// LS Electric XG5000 project: Trafic light3T
// PLC NewPLC
// module base 0 slot 0: Input/Output Module:XBM-DN32S (DC 24V INPUT/TR OUTPUT, 32points)
// module base 0 slot 1: Analog Input Module:XBF-AD04A (Volt/Current, 4-CH)
// module base 0 slot 2: Analog Output Module:XBF-DV04A (Voltage, 4-CH)

PROGRAM NewProgram (task: Scan Program)

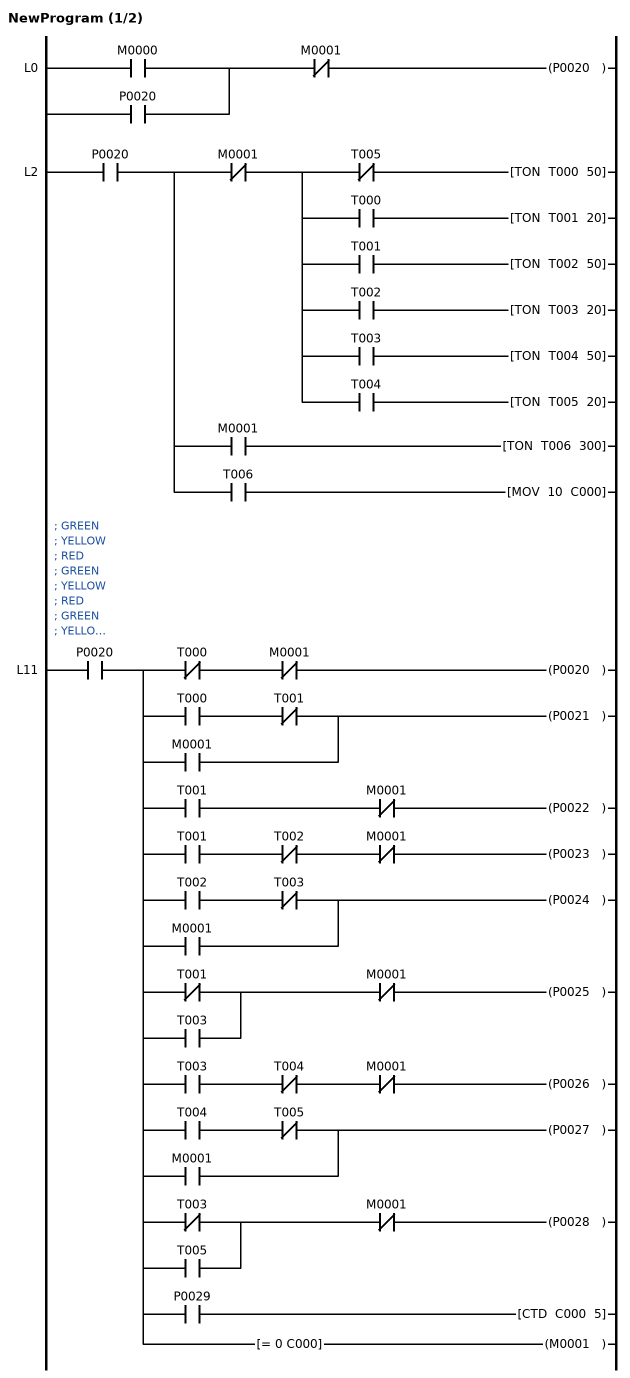
; L0
LOAD      M0000
OR        P0020
AND NOT   M0001
OUT       P0020
; L2
LOAD      P0020
MPUSH
AND NOT   M0001
MPUSH
AND NOT   T005
TON       T000 50
MLOAD
AND       T000
TON       T001 20
MLOAD
AND       T001
TON       T002 50
MLOAD
AND       T002
TON       T003 20
MLOAD
AND       T003
TON       T004 50
MPOP
AND       T004
TON       T005 20
MLOAD
AND       M0001
TON       T006 300
MPOP
AND       T006
MOV       10 C000
// output comment: 
; L11
LOAD      P0020
MPUSH
AND NOT   T000
AND NOT   M0001
OUT       P0020
MLOAD
LOAD      T000
AND NOT   T001
OR        M0001
AND LOAD
OUT       P0021
MLOAD
AND       T001
AND NOT   M0001
OUT       P0022
MLOAD
AND       T001
AND NOT   T002
AND NOT   M0001
OUT       P0023
MLOAD
LOAD      T002
AND NOT   T003
OR        M0001
AND LOAD
OUT       P0024
MLOAD
LOAD NOT  T001
OR        T003
AND LOAD
AND NOT   M0001
OUT       P0025
MLOAD
AND       T003
AND NOT   T004
AND NOT   M0001
OUT       P0026
MLOAD
LOAD      T004
AND NOT   T005
OR        M0001
AND LOAD
OUT       P0027
MLOAD
LOAD NOT  T003
OR        T005
AND LOAD
AND NOT   M0001
OUT       P0028
MLOAD
AND       P0029
CTD       C000 5
MPOP
AND=      0 C000
OUT       M0001
// output comment: GREEN 
// output comment: YELLOW
// output comment: RED
// output comment: GREEN 
// output comment: YELLOW
// output comment: RED
// output comment: GREEN
// output comment: YELLOW
// output comment: RED

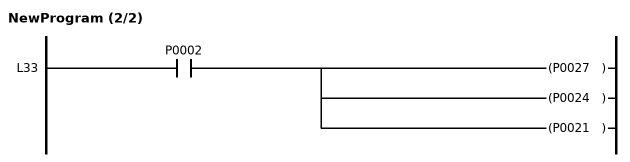
; L33
LOAD      P0002
OUT       P0027
OUT       P0024
OUT       P0021